FUNCTION_BLOCK AlarmesHabilitados (* Alarmes de limite do AnalogInput so quando habilitados (alarme desabilitado nao bloqueia nada) *)
  (* Standard: 61499-2 *)
  (* Version 1.1, 05/11/2026, Hidryco, Hidryco, 1.1: eventos de saida listados no ECAction (sem isso o runtime nao emite nenhum; o ST so liga/desliga). 1.0: saida = LimitReached AND NOT Disabled de cada alarme (HH, H, L, LL, ROC, DEV). O LimitReached da SE.App2Base compara mesmo com o alarme desabilitado. REQ recalcula e sempre emite CNF (mesmo tempo de hoje); REQ_DIS (mudanca de ajuste) so derruba os desabilitados e emite CNF se mudou. Usado no AnalogInput. *)
  PACKAGE SE.Nereda;
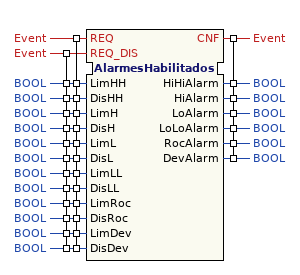
  EVENT_INPUT
    REQ WITH LimHH, DisHH, LimH, DisH, LimL, DisL, LimLL, DisLL, LimRoc, DisRoc, LimDev, DisDev; (* Novo estado dos alarmes (CNF dos alarmes) *)
    REQ_DIS WITH LimHH, DisHH, LimH, DisH, LimL, DisL, LimLL, DisLL, LimRoc, DisRoc, LimDev, DisDev; (* Ajuste ou habilitacao mudou (CNF_LIMITSP / IND dos alarmes) *)
  END_EVENT
  EVENT_OUTPUT
    CNF WITH HiHiAlarm, HiAlarm, LoAlarm, LoLoAlarm, RocAlarm, DevAlarm; (* Alarmes so com habilitacao *)
  END_EVENT
  VAR_INPUT
    LimHH : BOOL; (* LimitReached do alarme HH *)
    DisHH : BOOL; (* Disabled do alarme HH *)
    LimH : BOOL; (* LimitReached do alarme H *)
    DisH : BOOL; (* Disabled do alarme H *)
    LimL : BOOL; (* LimitReached do alarme L *)
    DisL : BOOL; (* Disabled do alarme L *)
    LimLL : BOOL; (* LimitReached do alarme LL *)
    DisLL : BOOL; (* Disabled do alarme LL *)
    LimRoc : BOOL; (* LimitReached do alarme Roc *)
    DisRoc : BOOL; (* Disabled do alarme Roc *)
    LimDev : BOOL; (* LimitReached do alarme Dev *)
    DisDev : BOOL; (* Disabled do alarme Dev *)
  END_VAR
  VAR_OUTPUT
    HiHiAlarm : BOOL; (* Alarme HH so com o alarme habilitado *)
    HiAlarm : BOOL; (* Alarme H so com o alarme habilitado *)
    LoAlarm : BOOL; (* Alarme L so com o alarme habilitado *)
    LoLoAlarm : BOOL; (* Alarme LL so com o alarme habilitado *)
    RocAlarm : BOOL; (* Alarme Roc so com o alarme habilitado *)
    DevAlarm : BOOL; (* Alarme Dev so com o alarme habilitado *)
  END_VAR
  VAR
    oldHiHiAlarm : BOOL;
    oldHiAlarm : BOOL;
    oldLoAlarm : BOOL;
    oldLoLoAlarm : BOOL;
    oldRocAlarm : BOOL;
    oldDevAlarm : BOOL;
  END_VAR
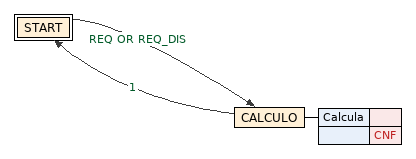
  EC_STATES
    START; (* Estado inicial *)
    CALCULO : Calcula, -> CNF; (* Calcula; o algoritmo decide se o CNF sai *)
  END_STATES
  EC_TRANSITIONS
    START TO CALCULO := REQ OR REQ_DIS;
    CALCULO TO START := 1;
  END_TRANSITIONS
  ALGORITHM Calcula IN ST: (* LimitReached AND NOT Disabled *)
CNF := FALSE;
IF REQ THEN
    (* mesmo momento de hoje: o CNF dos alarmes ja respeita o tempo do alarme *)
    HiHiAlarm := LimHH AND NOT DisHH;
    HiAlarm := LimH AND NOT DisH;
    LoAlarm := LimL AND NOT DisL;
    LoLoAlarm := LimLL AND NOT DisLL;
    RocAlarm := LimRoc AND NOT DisRoc;
    DevAlarm := LimDev AND NOT DisDev;
    CNF := TRUE;
ELSE
    (* mudanca de ajuste: so derruba quem foi desabilitado (habilitar espera o proximo CNF do alarme) *)
    HiHiAlarm := HiHiAlarm AND NOT DisHH;
    HiAlarm := HiAlarm AND NOT DisH;
    LoAlarm := LoAlarm AND NOT DisL;
    LoLoAlarm := LoLoAlarm AND NOT DisLL;
    RocAlarm := RocAlarm AND NOT DisRoc;
    DevAlarm := DevAlarm AND NOT DisDev;
    CNF := (HiHiAlarm <> oldHiHiAlarm) OR (HiAlarm <> oldHiAlarm) OR (LoAlarm <> oldLoAlarm) OR (LoLoAlarm <> oldLoLoAlarm) OR (RocAlarm <> oldRocAlarm) OR (DevAlarm <> oldDevAlarm);
END_IF;
oldHiHiAlarm := HiHiAlarm;
oldHiAlarm := HiAlarm;
oldLoAlarm := LoAlarm;
oldLoLoAlarm := LoLoAlarm;
oldRocAlarm := RocAlarm;
oldDevAlarm := DevAlarm;
  END_ALGORITHM
END_FUNCTION_BLOCK
